Universal Robots URScript: MAIN_1.script

# Set the default value
global current_frame, current_speed, current_acceleration, current_speedjoints, current_accelerationjoints, current_rounding
current_frame = [0.0, 0.0, 0.0, 0.0, 0.0, 0.0]
current_speed = 0.25
current_acceleration = 1.2
current_speedjoints = 1.0471975511965976
current_accelerationjoints = 1.3962634015954636
current_rounding = 0.0
#---------------------------------------------------------------------------------------------------------------------------
def MAIN_1():
  global current_instruction
# Program generated by RoboDK v5.6.9 for RoboDK Industrial on 26/02/2024 09:58:20
# Using nominal kinematics.
  current_instruction = "14: movej([-5.25645e-07, 0, 0, 0, 0, -1.46549e-15])"
  movej([-9.174235946645592e-09, 0.0, 0.0, 0.0, 0.0, -2.5577625655051703e-17],a=current_accelerationjoints,v=current_speedjoints,r=current_rounding)
  current_instruction = "16: movej([0, 3.21124, -15.4237, 0, 12.2125, -4.67269e-13])"
  movej([0.0, 0.05604671107174271, -0.2691943478398494, 0.0, 0.2131483348998075, -8.155382542501385e-15],a=current_accelerationjoints,v=current_speedjoints,r=current_rounding)
  current_instruction = "18: movel([1015, 0, 1272, 0.0, 90.0, 0.0])"
  movel(pose_trans(current_frame,[1.015000, 0.000000, 1.272000, 0.000000, 1.570796, 0.000000]),a=current_acceleration,v=current_speed,r=current_rounding)
  current_instruction = "20: setDO IO_Name:5 IO_Value:1"
  set_standard_digital_out(5,True)
  current_instruction = "22: waitDI IO_Name:5 IO_Value:1 Timeout(ms):-1"
  while True:
    sync()
    if get_standard_digital_in(5) == True:
      break
  end
  current_instruction = "28: waitDI IO_Name:5 IO_Value:1 Timeout(ms):100"
  myTimer = 0
  while True:
    myTimer = myTimer + get_steptime()
    sync()
    if myTimer >= 0.1:
      break
    if get_standard_digital_in(5) == True:
      break
  end
  popup(s='Message',title='Message',blocking=True)
  current_instruction = "39: 'REMOTE_PROG_CALL_171'"
  REMOTE_PROG_CALL_171()
  current_instruction = "41: 'CODE_INSERT_172'"
  CODE_INSERT_172
# Insert Comment
  global current_frame_name
  current_frame_name = 'Frame Pick and Place'
  global current_frame
  current_frame = [0.719013, -0.664003, 0.0, 0.0, 0.0, 0.0]
  global current_tcp
  current_tcp = [0.129073, 0.000000, 0.085477, 0.000000, 0.398790, 0.000000]
  set_tcp(current_tcp)
  global current_accelerationjoints
  current_accelerationjoints = 13.962634015954636
  global current_speedjoints
  current_speedjoints = 8.726646259971648
  global current_rounding
  current_rounding = 0.01
  current_instruction = "57: movej([-29.3322, 46.677, -0.024523, 26.5456, 25.3957, -51.634])"
  movej([-0.5119434668534807, 0.8146673349533932, -0.00042800709246656945, 0.4633081219174067, 0.443238580848724, -0.9011833059747522],a=current_accelerationjoints,v=current_speedjoints,r=current_rounding)
  global current_rounding
  current_rounding = -0.001
  global current_acceleration
  current_acceleration = 0.2
  global current_speed
  current_speed = 0.1
  current_instruction = "65: movel([187.786, 125.499, 139.112, 179.996, 0.18, -179.997])"
  movel(pose_trans(current_frame,[0.187786, 0.125499, 0.139112, 3.141523, 0.003142, -3.141540]),a=current_acceleration,v=current_speed,r=current_rounding)
  current_instruction = "67: setDO IO_Name:5 IO_Value:1"
  set_standard_digital_out(5,True)
  current_instruction = "69: 'PICK_PART_111'"
  PICK_PART_111()
  global current_rounding
  current_rounding = 0.01
  global current_acceleration
  current_acceleration = 0.6
  global current_speed
  current_speed = 0.3
# Linear movement using joint targets is not supported. Change the target type to cartesian or use a joint movement.
  current_instruction = "78: movel([187.272, 447.522, 305.347, -179.998, 0.18500000000000003, 179.999])"
  movel(pose_trans(current_frame,[0.187272, 0.447522, 0.305347, -3.141558, 0.003229, 3.141575]),a=current_acceleration,v=current_speed,r=current_rounding)
  global current_rounding
  current_rounding = -0.001
  global current_acceleration
  current_acceleration = 0.2
  global current_speed
  current_speed = 0.1
# MoveSearch command not implemented
  current_instruction = "87: movel([187.851, 447.517, 126.235, -179.998, 0.18500000000000003, 179.999])"
  movel(pose_trans(current_frame,[0.187851, 0.447517, 0.126235, -3.141558, 0.003229, 3.141575]),a=current_acceleration,v=current_speed,r=current_rounding)
  current_instruction = "89: setDO IO_Name:5 IO_Value:0"
  set_standard_digital_out(5,False)
  current_instruction = "91: 'PLACE_PART_112'"
  PLACE_PART_112()
  global current_rounding
  current_rounding = 0.01
  current_instruction = "95: movel([187.272, 447.522, 305.347, -179.998, 0.18500000000000003, 179.999])"
  movel(pose_trans(current_frame,[0.187272, 0.447522, 0.305347, -3.141558, 0.003229, 3.141575]),a=current_acceleration,v=current_speed,r=current_rounding)
  global current_frame_name
  current_frame_name = 'Frame Circular'
  global current_frame
  current_frame = [0.5776699999999999, 0.39225, 0.0, 0.0, 0.0, 0.679971549930731]
  global current_rounding
  current_rounding = 0.025
  global current_accelerationjoints
  current_accelerationjoints = 13.962634015954636
  global current_speedjoints
  current_speedjoints = 8.726646259971648
  global current_acceleration
  current_acceleration = 0.2
  global current_speed
  current_speed = 0.1
  current_instruction = "111: movej([52.186, 45.6758, 6.92, 66.7342, 19.9323, -92.73])"
  movej([0.9108175234457608, 0.797193098482426, 0.1207767842380076, 1.1647315136843999, 0.3478842624952658, -1.618443815374342],a=current_accelerationjoints,v=current_speedjoints,r=current_rounding)
  current_instruction = "113: movec([430.047, 43.774, 231.503, 178.913, 11.1813, -134.54900000000004],[109.688, -153.222, 161.073, 178.913, 11.1813, -134.54900000000004])"
  movec(pose_trans(current_frame,[0.430047, 0.043774, 0.231503, 3.122621, 0.195150, -2.348323]),pose_trans(current_frame,[0.109688, -0.153222, 0.161073, 3.122621, 0.195150, -2.348323]),a=current_acceleration,v=current_speed,r=current_rounding,mode=1)
# Circular movement using joint targets is not supported. Change the target type to cartesian or use a joint movement.
  global current_rounding
  current_rounding = -0.001
  global current_acceleration
  current_acceleration = 0.2
  global current_speed
  current_speed = 0.1
  current_instruction = "122: movel([312.208, 292.214, 255.156, 178.913, 11.1813, -134.54900000000004])"
  movel(pose_trans(current_frame,[0.312208, 0.292214, 0.255156, 3.122621, 0.195150, -2.348323]),a=current_acceleration,v=current_speed,r=current_rounding)
  current_instruction = "124: movej([-5.25645e-07, 0, 0, 0, 0, -1.46549e-15])"
  movej([-9.174235946645592e-09, 0.0, 0.0, 0.0, 0.0, -2.5577625655051703e-17],a=current_accelerationjoints,v=current_speedjoints,r=current_rounding)
  global current_frame_name
  current_frame_name = 'Frame Inspection'
  global current_frame
  current_frame = [0.0, 0.782714, 0.37761, 0.0, 0.0, 0.0]
  current_instruction = "130: movej([88.676, 29.6016, -6.42883, -1.98422, 49.4792, 4.54769])"
  movej([1.5476881674984917, 0.5166453838583535, -0.11220425055098705, -0.034631172083921885, 0.8635749512527783, 0.07937216386002093],a=current_accelerationjoints,v=current_speedjoints,r=current_rounding)
  current_instruction = "132: movel([19.898, 174.307, 19.008, -179.533, -5.425989999999999, -94.9281])"
  movel(pose_trans(current_frame,[0.019898, 0.174307, 0.019008, -3.133442, -0.094701, -1.656808]),a=current_acceleration,v=current_speed,r=current_rounding)
  current_instruction = "134: movel([378.402, 174.416, 18.997, -179.533, -5.425989999999999, -94.9281])"
  movel(pose_trans(current_frame,[0.378402, 0.174416, 0.018997, -3.133442, -0.094701, -1.656808]),a=current_acceleration,v=current_speed,r=current_rounding)
  current_instruction = "136: movel([380.996, 112.363, 34.882, -178.348, -18.1364, -95.2937])"
  movel(pose_trans(current_frame,[0.380996, 0.112363, 0.034882, -3.112760, -0.316540, -1.663189]),a=current_acceleration,v=current_speed,r=current_rounding)
  current_instruction = "138: movel([16.551, 114.359, 34.226, -178.348, -18.1364, -95.2937])"
  movel(pose_trans(current_frame,[0.016551, 0.114359, 0.034226, -3.112760, -0.316540, -1.663189]),a=current_acceleration,v=current_speed,r=current_rounding)
  current_instruction = "140: movel([26.434, 54.524, 46.072, 179.585, 4.348249999999999, -95.46080000000002])"
  movel(pose_trans(current_frame,[0.026434, 0.054524, 0.046072, 3.134350, 0.075891, -1.666105]),a=current_acceleration,v=current_speed,r=current_rounding)
  current_instruction = "142: movel([385.448, 48.05, 45.137, 178.913, 11.1809, -95.5904])"
  movel(pose_trans(current_frame,[0.385448, 0.048050, 0.045137, 3.122621, 0.195144, -1.668367]),a=current_acceleration,v=current_speed,r=current_rounding)
  current_instruction = "144: movel([385.448, -1.625, 295.251, 178.913, 11.1809, -95.5904])"
  movel(pose_trans(current_frame,[0.385448, -0.001625, 0.295251, 3.122621, 0.195144, -1.668367]),a=current_acceleration,v=current_speed,r=current_rounding)
  current_instruction = "146: movej([-5.25645e-07, 0, 0, 0, 0, -1.46549e-15])"
  movej([-9.174235946645592e-09, 0.0, 0.0, 0.0, 0.0, -2.5577625655051703e-17],a=current_accelerationjoints,v=current_speedjoints,r=current_rounding)
  current_instruction = "148: 'EVENT_PROG_START_101'"
  EVENT_PROG_START_101()
  global current_rounding
  current_rounding = 0.001
  global current_speed
  current_speed = 1.0
  global current_frame_name
  current_frame_name = 'Frame Inspection'
  global current_frame
  current_frame = [0.013637, -0.84008, 0.0, 0.0, 0.0, -1.5707963267948966]
# Show Tool 1
  current_instruction = "159: movej([-68.0903, 24.2019, 26.7855, 38.2134, 36.2017, -98.7964])"
  movej([-1.188399923670695, 0.4224028402384156, 0.4674951667929411, 0.6669496483816011, 0.6318388598192313, -1.7243224691173258],a=current_accelerationjoints,v=current_speedjoints,r=current_rounding)
  current_instruction = "161: 'EVENT_PATH_APPROACH_102'"
  EVENT_PATH_APPROACH_102()
  current_instruction = "163: movel([-49.895, 253.259, 319.999, -179.975, 0.353, -90.0])"
  movel(pose_trans(current_frame,[-0.049895, 0.253259, 0.319999, -3.141156, 0.006161, -1.570796]),a=current_acceleration,v=current_speed,r=current_rounding)
  current_instruction = "165: movel([0, 250, 270, -179.975, 0.353, -90.0])"
  movel(pose_trans(current_frame,[0.000000, 0.250000, 0.270000, -3.141156, 0.006161, -1.570796]),a=current_acceleration,v=current_speed,r=current_rounding)
  current_instruction = "167: 'EVENT_PATH_START_103'"
  EVENT_PATH_START_103()
  global current_speed
  current_speed = 0.05
  current_instruction = "171: movel([35.579, 247.455, 270, -179.92500000000004, 0.345, -90.0])"
  movel(pose_trans(current_frame,[0.035579, 0.247455, 0.270000, -3.140284, 0.006021, -1.570796]),a=current_acceleration,v=current_speed,r=current_rounding)
  current_instruction = "173: movel([70.433, 239.873, 270, -179.876, 0.330998, -89.999])"
  movel(pose_trans(current_frame,[0.070433, 0.239873, 0.270000, -3.139428, 0.005777, -1.570779]),a=current_acceleration,v=current_speed,r=current_rounding)
  current_instruction = "175: movel([103.854, 227.408, 270, -179.831, 0.3099970000000001, -89.999])"
  movel(pose_trans(current_frame,[0.103854, 0.227408, 0.270000, -3.138643, 0.005410, -1.570779]),a=current_acceleration,v=current_speed,r=current_rounding)
  current_instruction = "177: movel([135.16, 210.313, 270, -179.788, 0.282996, -89.999])"
  movel(pose_trans(current_frame,[0.135160, 0.210313, 0.270000, -3.137893, 0.004939, -1.570779]),a=current_acceleration,v=current_speed,r=current_rounding)
  current_instruction = "179: movel([163.715, 188.937, 270, -179.75000000000003, 0.24999599999999997, -89.999])"
  movel(pose_trans(current_frame,[0.163715, 0.188937, 0.270000, -3.137229, 0.004363, -1.570779]),a=current_acceleration,v=current_speed,r=current_rounding)
  current_instruction = "181: movel([188.937, 163.715, 270, -179.71700000000004, 0.211995, -89.999])"
  movel(pose_trans(current_frame,[0.188937, 0.163715, 0.270000, -3.136653, 0.003700, -1.570779]),a=current_acceleration,v=current_speed,r=current_rounding)
  current_instruction = "183: movel([210.313, 135.16, 270, -179.689, 0.169995, -89.999])"
  movel(pose_trans(current_frame,[0.210313, 0.135160, 0.270000, -3.136165, 0.002967, -1.570779]),a=current_acceleration,v=current_speed,r=current_rounding)
  current_instruction = "185: movel([227.408, 103.854, 270, -179.668, 0.12399399999999998, -89.999])"
  movel(pose_trans(current_frame,[0.227408, 0.103854, 0.270000, -3.135798, 0.002164, -1.570779]),a=current_acceleration,v=current_speed,r=current_rounding)
  current_instruction = "187: movel([239.873, 70.433, 270, -179.654, 0.075, -90.0])"
  movel(pose_trans(current_frame,[0.239873, 0.070433, 0.270000, -3.135554, 0.001309, -1.570796]),a=current_acceleration,v=current_speed,r=current_rounding)
  current_instruction = "189: movel([247.455, 35.579, 270, -179.647, 0.025, -90.0])"
  movel(pose_trans(current_frame,[0.247455, 0.035579, 0.270000, -3.135432, 0.000436, -1.570796]),a=current_acceleration,v=current_speed,r=current_rounding)
  current_instruction = "191: movel([250, 0, 270, -179.647, -0.025, -90.0])"
  movel(pose_trans(current_frame,[0.250000, 0.000000, 0.270000, -3.135432, -0.000436, -1.570796]),a=current_acceleration,v=current_speed,r=current_rounding)
  current_instruction = "193: movel([247.455, -35.579, 270, -179.654, -0.075, -90.0])"
  movel(pose_trans(current_frame,[0.247455, -0.035579, 0.270000, -3.135554, -0.001309, -1.570796]),a=current_acceleration,v=current_speed,r=current_rounding)
  current_instruction = "195: movel([239.873, -70.433, 270, -179.668, -0.12399399999999998, -90.001])"
  movel(pose_trans(current_frame,[0.239873, -0.070433, 0.270000, -3.135798, -0.002164, -1.570814]),a=current_acceleration,v=current_speed,r=current_rounding)
  current_instruction = "197: movel([227.408, -103.854, 270, -179.689, -0.169995, -90.001])"
  movel(pose_trans(current_frame,[0.227408, -0.103854, 0.270000, -3.136165, -0.002967, -1.570814]),a=current_acceleration,v=current_speed,r=current_rounding)
  current_instruction = "199: movel([210.313, -135.16, 270, -179.71700000000004, -0.211995, -90.001])"
  movel(pose_trans(current_frame,[0.210313, -0.135160, 0.270000, -3.136653, -0.003700, -1.570814]),a=current_acceleration,v=current_speed,r=current_rounding)
  current_instruction = "201: movel([188.937, -163.715, 270, -179.75000000000003, -0.24999599999999997, -90.001])"
  movel(pose_trans(current_frame,[0.188937, -0.163715, 0.270000, -3.137229, -0.004363, -1.570814]),a=current_acceleration,v=current_speed,r=current_rounding)
  current_instruction = "203: movel([163.715, -188.937, 270, -179.788, -0.282996, -90.001])"
  movel(pose_trans(current_frame,[0.163715, -0.188937, 0.270000, -3.137893, -0.004939, -1.570814]),a=current_acceleration,v=current_speed,r=current_rounding)
  current_instruction = "205: movel([135.16, -210.313, 270, -179.83, -0.3109970000000001, -90.001])"
  movel(pose_trans(current_frame,[0.135160, -0.210313, 0.270000, -3.138626, -0.005428, -1.570814]),a=current_acceleration,v=current_speed,r=current_rounding)
  current_instruction = "207: movel([103.854, -227.408, 270, -179.876, -0.331998, -90.001])"
  movel(pose_trans(current_frame,[0.103854, -0.227408, 0.270000, -3.139428, -0.005794, -1.570814]),a=current_acceleration,v=current_speed,r=current_rounding)
  current_instruction = "209: movel([70.433, -239.873, 270, -179.92500000000004, -0.346, -90.0])"
  movel(pose_trans(current_frame,[0.070433, -0.239873, 0.270000, -3.140284, -0.006039, -1.570796]),a=current_acceleration,v=current_speed,r=current_rounding)
  current_instruction = "211: movel([35.579, -247.455, 270, -179.975, -0.353, -90.0])"
  movel(pose_trans(current_frame,[0.035579, -0.247455, 0.270000, -3.141156, -0.006161, -1.570796]),a=current_acceleration,v=current_speed,r=current_rounding)
  current_instruction = "213: movel([0, -250, 270, -179.975, -0.353, -90.0])"
  movel(pose_trans(current_frame,[0.000000, -0.250000, 0.270000, -3.141156, -0.006161, -1.570796]),a=current_acceleration,v=current_speed,r=current_rounding)
  current_instruction = "215: movel([0, -250, 270, 179.975, -0.353, -90.0])"
  movel(pose_trans(current_frame,[0.000000, -0.250000, 0.270000, 3.141156, -0.006161, -1.570796]),a=current_acceleration,v=current_speed,r=current_rounding)
  current_instruction = "217: movel([-35.579, -247.455, 270, 179.92500000000004, -0.346, -90.0])"
  movel(pose_trans(current_frame,[-0.035579, -0.247455, 0.270000, 3.140284, -0.006039, -1.570796]),a=current_acceleration,v=current_speed,r=current_rounding)
  current_instruction = "219: movel([-70.433, -239.873, 270, 179.876, -0.330998, -89.999])"
  movel(pose_trans(current_frame,[-0.070433, -0.239873, 0.270000, 3.139428, -0.005777, -1.570779]),a=current_acceleration,v=current_speed,r=current_rounding)
  current_instruction = "221: movel([-103.854, -227.408, 270, 179.831, -0.3099970000000001, -89.999])"
  movel(pose_trans(current_frame,[-0.103854, -0.227408, 0.270000, 3.138643, -0.005410, -1.570779]),a=current_acceleration,v=current_speed,r=current_rounding)
  current_instruction = "223: movel([-135.16, -210.313, 270, 179.788, -0.282996, -89.999])"
  movel(pose_trans(current_frame,[-0.135160, -0.210313, 0.270000, 3.137893, -0.004939, -1.570779]),a=current_acceleration,v=current_speed,r=current_rounding)
  current_instruction = "225: movel([-163.715, -188.937, 270, 179.75000000000003, -0.24999599999999997, -89.999])"
  movel(pose_trans(current_frame,[-0.163715, -0.188937, 0.270000, 3.137229, -0.004363, -1.570779]),a=current_acceleration,v=current_speed,r=current_rounding)
  current_instruction = "227: movel([-188.937, -163.715, 270, 179.71700000000004, -0.211995, -89.999])"
  movel(pose_trans(current_frame,[-0.188937, -0.163715, 0.270000, 3.136653, -0.003700, -1.570779]),a=current_acceleration,v=current_speed,r=current_rounding)
  current_instruction = "229: movel([-210.313, -135.16, 270, 179.69, -0.168995, -89.999])"
  movel(pose_trans(current_frame,[-0.210313, -0.135160, 0.270000, 3.136182, -0.002950, -1.570779]),a=current_acceleration,v=current_speed,r=current_rounding)
  current_instruction = "231: movel([-227.408, -103.854, 270, 179.669, -0.12299400000000002, -89.999])"
  movel(pose_trans(current_frame,[-0.227408, -0.103854, 0.270000, 3.135816, -0.002147, -1.570779]),a=current_acceleration,v=current_speed,r=current_rounding)
  current_instruction = "233: movel([-239.873, -70.433, 270, 179.654, -0.075, -90.0])"
  movel(pose_trans(current_frame,[-0.239873, -0.070433, 0.270000, 3.135554, -0.001309, -1.570796]),a=current_acceleration,v=current_speed,r=current_rounding)
  current_instruction = "235: movel([-247.455, -35.579, 270, 179.647, -0.025, -90.0])"
  movel(pose_trans(current_frame,[-0.247455, -0.035579, 0.270000, 3.135432, -0.000436, -1.570796]),a=current_acceleration,v=current_speed,r=current_rounding)
  current_instruction = "237: movel([-250, 0, 270, 179.647, 0.025, -90.0])"
  movel(pose_trans(current_frame,[-0.250000, 0.000000, 0.270000, 3.135432, 0.000436, -1.570796]),a=current_acceleration,v=current_speed,r=current_rounding)
  current_instruction = "239: movel([-247.455, 35.579, 270, 179.655, 0.075, -90.0])"
  movel(pose_trans(current_frame,[-0.247455, 0.035579, 0.270000, 3.135571, 0.001309, -1.570796]),a=current_acceleration,v=current_speed,r=current_rounding)
  current_instruction = "241: movel([-239.873, 70.433, 270, 179.669, 0.12299400000000002, -90.001])"
  movel(pose_trans(current_frame,[-0.239873, 0.070433, 0.270000, 3.135816, 0.002147, -1.570814]),a=current_acceleration,v=current_speed,r=current_rounding)
  current_instruction = "243: movel([-227.408, 103.854, 270, 179.689, 0.169995, -90.001])"
  movel(pose_trans(current_frame,[-0.227408, 0.103854, 0.270000, 3.136165, 0.002967, -1.570814]),a=current_acceleration,v=current_speed,r=current_rounding)
  current_instruction = "245: movel([-210.313, 135.16, 270, 179.71700000000004, 0.211995, -90.001])"
  movel(pose_trans(current_frame,[-0.210313, 0.135160, 0.270000, 3.136653, 0.003700, -1.570814]),a=current_acceleration,v=current_speed,r=current_rounding)
  current_instruction = "247: movel([-188.937, 163.715, 270, 179.75000000000003, 0.24999599999999997, -90.001])"
  movel(pose_trans(current_frame,[-0.188937, 0.163715, 0.270000, 3.137229, 0.004363, -1.570814]),a=current_acceleration,v=current_speed,r=current_rounding)
  current_instruction = "249: movel([-163.715, 188.937, 270, 179.788, 0.282996, -90.001])"
  movel(pose_trans(current_frame,[-0.163715, 0.188937, 0.270000, 3.137893, 0.004939, -1.570814]),a=current_acceleration,v=current_speed,r=current_rounding)
  current_instruction = "251: movel([-135.16, 210.313, 270, 179.831, 0.3099970000000001, -90.001])"
  movel(pose_trans(current_frame,[-0.135160, 0.210313, 0.270000, 3.138643, 0.005410, -1.570814]),a=current_acceleration,v=current_speed,r=current_rounding)
  current_instruction = "253: movel([-103.854, 227.408, 270, 179.876, 0.331998, -90.001])"
  movel(pose_trans(current_frame,[-0.103854, 0.227408, 0.270000, 3.139428, 0.005794, -1.570814]),a=current_acceleration,v=current_speed,r=current_rounding)
  current_instruction = "255: movel([-70.433, 239.873, 270, 179.92500000000004, 0.346, -90.0])"
  movel(pose_trans(current_frame,[-0.070433, 0.239873, 0.270000, 3.140284, 0.006039, -1.570796]),a=current_acceleration,v=current_speed,r=current_rounding)
  current_instruction = "257: movel([-35.579, 247.455, 270, 179.975, 0.353, -90.0])"
  movel(pose_trans(current_frame,[-0.035579, 0.247455, 0.270000, 3.141156, 0.006161, -1.570796]),a=current_acceleration,v=current_speed,r=current_rounding)
  current_instruction = "259: movel([0, 250, 270, 179.975, 0.353, -90.0])"
  movel(pose_trans(current_frame,[0.000000, 0.250000, 0.270000, 3.141156, 0.006161, -1.570796]),a=current_acceleration,v=current_speed,r=current_rounding)
  global current_speed
  current_speed = 1.0
  current_instruction = "263: 'EVENT_PATH_FINISH_105'"
  EVENT_PATH_FINISH_105()
  current_instruction = "265: movel([49.895, 253.258, 319.999, 179.975, 0.353, -90.0])"
  movel(pose_trans(current_frame,[0.049895, 0.253258, 0.319999, 3.141156, 0.006161, -1.570796]),a=current_acceleration,v=current_speed,r=current_rounding)
  current_instruction = "267: movel([49.939, 252.642, 419.997, 179.975, 0.353, -90.0])"
  movel(pose_trans(current_frame,[0.049939, 0.252642, 0.419997, 3.141156, 0.006161, -1.570796]),a=current_acceleration,v=current_speed,r=current_rounding)
  current_instruction = "269: 'EVENT_PATH_RETRACT_106'"
  EVENT_PATH_RETRACT_106()
  current_instruction = "271: 'EVENT_PROG_FINISH_107'"
  EVENT_PROG_FINISH_107()
  global current_frame_name
  current_frame_name = 'Frame Pick and Place'
  global current_frame
  current_frame = [0.719013, -0.664003, 0.0, 0.0, 0.0, 0.0]
  current_instruction = "277: movej([-29.3322, 46.677, -0.024523, 26.5456, 25.3957, -51.634])"
  movej([-0.5119434668534807, 0.8146673349533932, -0.00042800709246656945, 0.4633081219174067, 0.443238580848724, -0.9011833059747522],a=current_accelerationjoints,v=current_speedjoints,r=current_rounding)
  current_instruction = "279: sleep(1250.0ms)"
  sleep(1.25)
  current_instruction = "281: movel([187.786, 125.499, 139.112, 179.996, 0.18, -179.997])"
  movel(pose_trans(current_frame,[0.187786, 0.125499, 0.139112, 3.141523, 0.003142, -3.141540]),a=current_acceleration,v=current_speed,r=current_rounding)
  current_instruction = "283: waitDI IO_Name:1 IO_Value:1 Timeout(ms):-1"
  while True:
    sync()
    if get_standard_digital_in(1) == True:
      break
  end
  current_instruction = "289: movel([187.264, 125.487, 305.356, -180.0, 0.184, 180.0])"
  movel(pose_trans(current_frame,[0.187264, 0.125487, 0.305356, -3.141593, 0.003211, 3.141593]),a=current_acceleration,v=current_speed,r=current_rounding)
  current_instruction = "291: 'PROG 1 _.-[]/\\;,><&*:%=+@!#^|?^ with a very long name and special characters'"
  PROG_1__________________________with_a_very_long_name_and_special_characters()
end
def PROG_1__________________________with_a_very_long_name_and_special_characters():
  global current_instruction
# This is a subprogram call to PROG_1
  global current_frame_name
  current_frame_name = 'Frame 1 _.-[]/\\;,><&*:%=+@!#^|?^ with a very long name and special characters'
  global current_frame
  current_frame = [0.0, 1.0, 0.0, 0.0, 0.0, 0.0]
  global current_tcp
  current_tcp = [0.000000, 0.000000, 0.200000, 0.000000, 0.000000, 0.000000]
  set_tcp(current_tcp)
  current_instruction = "304: movej([-5.25645e-07, 0, 0, 0, 0, -3.50835e-15])"
  movej([-9.174235946645592e-09, 0.0, 0.0, 0.0, 0.0, -6.123225881234306e-17],a=current_accelerationjoints,v=current_speedjoints,r=current_rounding)
end
MAIN_1()
